// The IAG50cm telescope on mock axes, scanned in the MAIN order (axes, then the telescope; IAG50cm/POUs/MAIN.TcPOU).
// One Scan() is one PLC scan. The scenario tests own one rig each (VAR_INST of the test method) and call Scan() once per
// PLC cycle: the astronomical clock needs a real NT_GetTime round trip (up to about 5 s) before FB_TelescopeControl accepts a
// goto/slew/track, so a rig is not usable before ClockValid. Everything else counts scans, not time.
// Plan: BROTLib specs/plans/2026-10-21-telescope-state-machine-unification.md (D1, step 2).
FUNCTION_BLOCK FB_IagRig
VAR
	fbComm			: FB_RecordingComm;	// records nothing until a test calls Start (IagTelemetry_Tests)
	fbHa			: FB_HourAngleMock(comm := fbComm);
	fbDec			: FB_DeclinationMock(comm := fbComm);
	fbFocus			: FB_FocusMock;
	fbCovers		: FB_CoversMock;
	fbDome			: FB_DomeMock;
	fbTel			: FB_TelescopeControl(comm := fbComm);
	pBool			: POINTER TO BOOL;
	nScans			: UDINT;
	nTimeDivisor	: UDINT := 1;	// the time seam of the telescope under test (SetTimeDivisor)
	fHorizon		: LREAL := 1.0;	// the horizon limit passed to the telescope (an input, so tests set it here; #84)
END_VAR
VAR CONSTANT
	telescopeConfig	: ST_TelescopeConfig := (longitude := 9.9452433, latitude := 51.5592378, altitude := 100.0,
											 houranglePark := 0.0, declinationPark := 52.0, focusPark := 16.3,
											 hourangleHome := 0.0, declinationHome := 52.0, focusHome := 16.3,
											 name := 'Emmy Noether', diameter := 0.5, cabinet := 'Beckhoff', manufacturer := 'test',
											 mountOptions := 'HA-DEC', mount := 'HA_DEC');
END_VAR

METHOD Scan
// the five contacts the cabinet error is made of (FB_CabinetControl, #10); unlinked they read FALSE
pBool := ADR(fbTel.fbCabinet.bAuxiliaryContact24V);		pBool^ := TRUE;
pBool := ADR(fbTel.fbCabinet.bAuxiliaryContact48V);		pBool^ := TRUE;
pBool := ADR(fbTel.fbCabinet.bAuxiliaryContactHADEC);	pBool^ := TRUE;
pBool := ADR(fbTel.fbCabinet.bAuxiliaryContactFOCUS);	pBool^ := TRUE;
pBool := ADR(fbTel.fbCabinet.bCollectiveReport24VFuse);	pBool^ := TRUE;

fbHa();
fbDec();
fbFocus();
fbTel(
	fbHourAngle := fbHa,
	fbDeclination := fbDec,
	fbFocus := fbFocus,
	fbDome := fbDome,
	fbCovers := fbCovers,
	telescopeConfig := telescopeConfig,
	nTimeDivisor := nTimeDivisor,
	fHorizon := fHorizon);
nScans := nScans + 1;
END_METHOD

PROPERTY ClockValid : BOOL
GET
ClockValid := fbTel.fbTime.bValid;
END_GET
END_PROPERTY

PROPERTY Online : BOOL
GET
Online := fbTel.ReadyState = 1.0;
END_GET
END_PROPERTY

// divides every long timeout of the telescope (600 s, 2 min, 12 h) by nValue, for this rig only (1 = real times)
METHOD SetTimeDivisor
VAR_INPUT
	nValue	: UDINT;
END_VAR
nTimeDivisor := nValue;
fbTel.nTimeDivisor := nValue;
END_METHOD

// the horizon limit of the telescope under test (an input of the telescope, so it cannot be written from outside; #84)
METHOD SetHorizon
VAR_INPUT
	fValue	: LREAL;
END_VAR
fHorizon := fValue;
END_METHOD

// scans a move takes on both mock axes (default 60)
METHOD SetMoveScans
VAR_INPUT
	nScans	: UINT;
END_VAR
fbHa.nMockMoveScans := nScans;
fbDec.nMockMoveScans := nScans;
END_METHOD

// scans the calibration sweep (homing) of each mock axis takes (default 3, #197)
METHOD SetHomeScans
VAR_INPUT
	nHa		: UINT;
	nDec	: UINT;
END_VAR
fbHa.nMockHomeScans := nHa;
fbDec.nMockHomeScans := nDec;
END_METHOD

// scans from a move command until the mock axes report InMotion (default 0: at once); the NC on the real axes takes a few cycles
METHOD SetStartScans
VAR_INPUT
	nScans	: UINT;
END_VAR
fbHa.nMockStartScans := nScans;
fbDec.nMockStartScans := nScans;
END_METHOD

// #120: the stop of the mock axis ends at rest but never reports Done (a lost Done, or a stop that was never allowed)
METHOD SetStopWithoutDone
VAR_INPUT
	bHa		: BOOL;
	bDec	: BOOL;
END_VAR
fbHa.bMockNoStopDone := bHa;
fbDec.bMockNoStopDone := bDec;
END_METHOD

// the user offsets of the telescope under test (degrees; IAG50cm#17 telemetry tests)
METHOD SetOffsets
VAR_INPUT
	fHourAngle	: LREAL;
	fDeclination	: LREAL;
END_VAR
fbTel.HourAngleOffset := fHourAngle;
fbTel.DeclinationOffset := fDeclination;
END_METHOD

// the command input bStop of the telescope under test, as an ADS writer sets it (not the method)
METHOD SetStopInput
VAR_INPUT
	bValue	: BOOL;
END_VAR
fbTel.bStop := bValue;
END_METHOD

// the command input bPark of the telescope under test, as an ADS writer sets it (not the method)
METHOD SetParkInput
VAR_INPUT
	bValue	: BOOL;
END_VAR
fbTel.bPark := bValue;
END_METHOD

// the command input bPower of the telescope under test, as an ADS writer sets it (not the method)
METHOD SetPowerInput
VAR_INPUT
	bValue	: BOOL;
END_VAR
fbTel.bPower := bValue;
END_METHOD

// the command input bSlew of the telescope under test, as an ADS writer sets it (not the method)
METHOD SetSlewInput
VAR_INPUT
	bValue	: BOOL;
END_VAR
fbTel.bSlew := bValue;
END_METHOD

// the slew target fields an ADS writer sets before it raises bSlew
METHOD SetSlewTargetInput
VAR_INPUT
	fAzimuth	: LREAL;
	fAltitude	: LREAL;
END_VAR
fbTel.fAzimuth := fAzimuth;
fbTel.fElevation := fAltitude;
END_METHOD

// the command input bTrack of the telescope under test, as an ADS writer sets it (not the method)
METHOD SetTrackInput
VAR_INPUT
	bValue	: BOOL;
END_VAR
fbTel.bTrack := bValue;
END_METHOD

// sets the request latch bGoHomeActive of the telescope under test (an output, written through a pointer): a request left over from before

METHOD ForceGoHomeActive
pBool := ADR(fbTel.bGoHomeActive);

pBool^ := TRUE;
END_METHOD

// sets the request latch bSlewActive of the telescope under test (an output, written through a pointer): a request left over from before

METHOD ForceSlewActive
pBool := ADR(fbTel.bSlewActive);

pBool^ := TRUE;
END_METHOD

// the pointing-model safe altitude of the telescope under test (an input of the telescope; a goto target below it is refused)

METHOD SetSafeAltitude

VAR_INPUT

	fValue	: LREAL;

END_VAR
fbTel.fPointingSafeAltitude := fValue;
END_METHOD

// the E-stop input of the telescope under test (#14)
METHOD SetEstop
VAR_INPUT
	bValue	: BOOL;
END_VAR
fbTel.bEstopTriggered := bValue;
END_METHOD

METHOD InjectHaError
VAR_INPUT
	nId	: UDINT;
END_VAR
fbHa.InjectError(nId);
END_METHOD

METHOD InjectDecError
VAR_INPUT
	nId	: UDINT;
END_VAR
fbDec.InjectError(nId);
END_METHOD

END_FUNCTION_BLOCK

(* stored: Version 1.1.0.1, ProductVersion 3.1.4024.15
   POU FB_IagRig: Id {f911297a-7486-47f1-9f44-b3154b341e1d}, SpecialFunc None
   Method Scan: Id {fa6422ce-24fd-4aeb-b8a7-2d38ea6a1e96}
   Property ClockValid: Id {a65ae0e9-65c9-4b55-8f9e-7139e8ee047a}
   Get Get: Id {b2e5b616-98ac-4ad2-8d2b-76302ac69731}
   Property Online: Id {dbe83508-7e2e-403f-9bf0-c4cf26a65310}
   Get Get: Id {69a3b469-7b54-4fd0-894e-68b9927ea365}
   Method SetTimeDivisor: Id {26d99b39-b426-4fd5-ac43-ba739ce53716}
   Method SetHorizon: Id {40095ef5-bf79-47cb-b27f-9ceb704f18d1}
   Method SetMoveScans: Id {cdeb9136-db3d-432e-8efa-7f4fddc23765}
   Method SetHomeScans: Id {3b8e5d17-6a42-4c90-8f1d-72e4a0c9b315}
   Method SetStartScans: Id {933a0b2d-7791-43fd-bb42-99ec4e6a5ddf}
   Method SetStopWithoutDone: Id {31dd82bd-7635-43b2-809d-d1cf60884bb0}
   Method SetOffsets: Id {7c1d4a52-3be0-4f0b-9a5e-0d6a1c2f8b11}
   Method SetStopInput: Id {7bdbc188-a661-4e04-b5d2-f62e1fdab845}
   Method SetParkInput: Id {28ebb24d-6560-49cd-8361-4560c35e2adc}
   Method SetPowerInput: Id {32f6aaab-4cad-4b81-b9f1-72e3e4955e55}
   Method SetSlewInput: Id {56f9b5ac-d946-4b7f-bf1f-220a8f105ee7}
   Method SetSlewTargetInput: Id {5fe36a9f-ab27-440f-842f-bdba6e7ceba4}
   Method SetTrackInput: Id {5afafdc8-4a81-4113-9b6a-42ca03f9727f}
   Method ForceGoHomeActive: Id {abb77387-5b6c-4636-bc8b-2a95b777a604}
   Method ForceSlewActive: Id {3ffb04e7-864e-4540-994d-94252b727107}
   Method SetSafeAltitude: Id {5080fecd-12c1-4a4d-85b0-db08c61b38f5}
   Method SetEstop: Id {2e9b6f03-51a7-4c8d-b3f4-8a7d90e1c622}
   Method InjectHaError: Id {905dc23c-55b4-4eb7-a513-f6b52cccde02}
   Method InjectDecError: Id {1a4cba55-34b7-4db9-ad88-e6e39d342843} *)
